(* IEC 61131-3 sources: SRCI_CLIENT_PLC/RobotLibrary/Library/POUs/BasicMove/MC_ReturnToPrimary/Structures, 4 files *)

(* ---- ReturnToPrimaryOutCmd.st ---- *)
{attribute 'pack_mode' := '1'}
// -------------------------------------------------------------------------
//  SRCI Robot Library
// -------------------------------------------------------------------------
//
//  Object:      ReturnToPrimaryOutCmd
//  Author:      Thorsten Brach
//  Date:        2024-06-22
//
//  Description:
//
//
//  Copyright:
//    (C) 2024 Thorsten Brach. All rights reserved
//             Licensed under the MIT License.
//
//  Disclaimer:
//    This project is provided without any guarantee and can be used for
//    private and commercial purposes. Any use is at the user’s
//    own risk and responsibility.
//
// -------------------------------------------------------------------------
TYPE ReturnToPrimaryOutCmd :
STRUCT
  /// Distance-to-go of the current job.
  /// • -1: No valid value because move command is not yet active (valid values are pending) or not supported by RC
  /// • >0: Actual distance between current and target position
  /// •  0: Target position reached
  RemainingDistance  : REAL;
  /// Percentage of already traversed distance of current job.
  /// If not supported : • -1
  Progress           : REAL;
  /// Tool index of target position of ReturnToPrimary
  /// • 0: Flange
  /// • 1..254: Tool frames
  PrimaryPosToolNo   : USINT;
  /// Frame index of target position of ReturnToPrimary
  /// • 0: WCS
  ///• 1..254: User frames
  PrimaryPosFrameNo  : USINT;
END_STRUCT
END_TYPE

(* ---- ReturnToPrimaryParCmd.st ---- *)
{attribute 'pack_mode' := '1'}
// -------------------------------------------------------------------------
//  SRCI Robot Library
// -------------------------------------------------------------------------
//
//  Object:      ReturnToPrimaryParCmd
//  Author:      Thorsten Brach
//  Date:        2024-06-22
//
//  Description:
//
//
//  Copyright:
//    (C) 2024 Thorsten Brach. All rights reserved
//             Licensed under the MIT License.
//
//  Disclaimer:
//    This project is provided without any guarantee and can be used for
//    private and commercial purposes. Any use is at the user’s
//    own risk and responsibility.
//
// -------------------------------------------------------------------------
TYPE ReturnToPrimaryParCmd :
STRUCT
  /// Defines target position when function is executed:
  /// • 0: Interrupt position (default) - Returns to position active,  when interrupt was executed
  /// • 1: End position                 - Returns to target position of interrupted segment
  ReturnMode         : ReturnMode;
  /// TCP velocity in % of nominal velocity
  /// •  <0%: (default) - Use default velocity
  /// •   0%:           - Use internal minimal velocity
  /// • 100%:           - Use maximal reference velocity
  /// See chapter 5.5.7 Robot dynamics
  VelocityRate       : REAL := -1.0; // ST-FIX F41: spec 5.x robot dynamics parameter: '<0 %: use default' (default); the library had 0.0 = internal minimal value (the RC rejects 0 for DecelerationRate/JerkRate)
  /// Acceleration for movement in % of nominal acceleration
  /// •  <0%: (default) - Use default acceleration
  /// •   0%:           - Use internal minimal acceleration
  /// • 100%:           - Use maximal reference acceleration
  /// See chapter 5.5.7 Robot dynamics
  AccelerationRate   : REAL := -1.0; // ST-FIX F41: spec 5.x robot dynamics parameter: '<0 %: use default' (default); the library had 0.0 = internal minimal value (the RC rejects 0 for DecelerationRate/JerkRate)
  /// Deceleration for movement in % of nominal deceleration
  /// •  <0%: (default) - Use default deceleration
  /// •   0%:           - Use internal minimal deceleration
  /// • 100%:           - Use maximal reference deceleration
  /// See chapter 5.5.7 Robot dynamics
  DecelerationRate   : REAL := -1.0; // ST-FIX F41: spec 5.x robot dynamics parameter: '<0 %: use default' (default); the library had 0.0 = internal minimal value (the RC rejects 0 for DecelerationRate/JerkRate)
  /// Jerk of the movement in % of nominal jerk
  /// •  <0%: (default) - Use default jerk
  /// •   0%:           - Use internal minimal jerk
  /// • 100%:           - Use maximal reference jerk
  /// See chapter 5.5.7 Robot dynamics
  JerkRate           : REAL := -1.0; // ST-FIX F41: spec 5.x robot dynamics parameter: '<0 %: use default' (default); the library had 0.0 = internal minimal value (the RC rejects 0 for DecelerationRate/JerkRate)
  /// Index of tool
  /// •      0: Flange (default)
  /// • 1..254: Tool frames
  ToolNo             : USINT;
  /// Index of frame
  /// •      0: WCS (default)
  /// • 1..254: User frames
  FrameNo            : USINT;
  /// Parameter is used if it is greater than 0 (default):
  /// Maximum allowed distance between current position and target position according to ReturnMode.
  /// If calculated distance is beyond specified Limit, RC returns an error
  DistanceLimit      : REAL;
  /// Defines type of command movement. One of the optional modes must be supported
  TrajectoryMode     : TrajectoryMode;
  /// Parameter is used if it is greater than 0 (default)
  /// • Velocity input is ignored
  /// • Parameter defines the time for the movement to reach the target position
  /// Error is sent by the RC if the time cannot be kept
  MoveTime           : TIME;
  /// Set TRUE to deactivate comparison of
  /// • ToolData and FrameData
  /// • ToolNo and PrimaryPosToolNo
  /// • FrameNo and PrimaryPosFrameNo
  AllowDifferences   : BOOL;
END_STRUCT
END_TYPE

(* ---- ReturnToPrimaryRecvData.st ---- *)
{attribute 'pack_mode' := '1'}
// -------------------------------------------------------------------------
//  SRCI Robot Library
// -------------------------------------------------------------------------
//
//  Object:      ReturnToPrimaryRecvData
//  Author:      Thorsten Brach
//  Date:        2024-06-22
//
//  Description:
//
//
//  Copyright:
//    (C) 2024 Thorsten Brach. All rights reserved
//             Licensed under the MIT License.
//
//  Disclaimer:
//    This project is provided without any guarantee and can be used for
//    private and commercial purposes. Any use is at the user’s
//    own risk and responsibility.
//
// -------------------------------------------------------------------------
TYPE ReturnToPrimaryRecvData EXTENDS RspHeader :
STRUCT
  /// Percentage of already traversed distance of current job.
  /// If not supported : • -1
  Progress           : UINT;
  /// Distance-to-go of the current job.
  /// • -1: No valid value because move command is not yet active (valid values are pending) or not supported by RC
  /// • >0: Actual distance between current and target position
  /// •  0: Target position reached
  RemainingDistance  : REAL;
  /// Tool index of target position of ReturnToPrimary
  /// • 0: Flange
  /// • 1..254: Tool frames
  PrimaryPosToolNo   : USINT;
  /// Frame index of target position of ReturnToPrimary
  /// • 0: WCS
  ///• 1..254: User frames
  PrimaryPosFrameNo  : USINT;
END_STRUCT
END_TYPE

(* ---- ReturnToPrimarySendData.st ---- *)
{attribute 'pack_mode' := '1'}
// -------------------------------------------------------------------------
//  SRCI Robot Library
// -------------------------------------------------------------------------
//
//  Object:      ReturnToPrimarySendData
//  Author:      Thorsten Brach
//  Date:        2024-06-22
//
//  Description:
//
//
//  Copyright:
//    (C) 2024 Thorsten Brach. All rights reserved
//             Licensed under the MIT License.
//
//  Disclaimer:
//    This project is provided without any guarantee and can be used for
//    private and commercial purposes. Any use is at the user’s
//    own risk and responsibility.
//
// -------------------------------------------------------------------------
TYPE ReturnToPrimarySendData EXTENDS CmdHeader:
STRUCT
  /// TCP velocity in % of nominal velocity
  /// •  <0%: (default) - Use default velocity
  /// •   0%:           - Use internal minimal velocity
  /// • 100%:           - Use maximal reference velocity
  /// See chapter 5.5.7 Robot dynamics
  VelocityRate       : UINT;
  /// Acceleration for movement in % of nominal acceleration
  /// •  <0%: (default) - Use default acceleration
  /// •   0%:           - Use internal minimal acceleration
  /// • 100%:           - Use maximal reference acceleration
  /// See chapter 5.5.7 Robot dynamics
  AccelerationRate   : UINT;
  /// Deceleration for movement in % of nominal deceleration
  /// •  <0%: (default) - Use default deceleration
  /// •   0%:           - Use internal minimal deceleration
  /// • 100%:           - Use maximal reference deceleration
  /// See chapter 5.5.7 Robot dynamics
  DecelerationRate   : UINT;
  /// Jerk of the movement in % of nominal jerk
  /// •  <0%: (default) - Use default jerk
  /// •   0%:           - Use internal minimal jerk
  /// • 100%:           - Use maximal reference jerk
  /// See chapter 5.5.7 Robot dynamics
  JerkRate           : UINT;
  /// Parameter is used if it is greater than 0 (default):
  /// Maximum allowed distance between current position and target position according to ReturnMode.
  /// If calculated distance is beyond specified Limit, RC returns an error
  DistanceLimit      : REAL;
  /// Index of tool
  /// •      0: Flange (default)
  /// • 1..254: Tool frames
  ToolNo             : USINT;
  /// Index of frame
  /// •      0: WCS (default)
  /// • 1..254: User frames
  FrameNo            : USINT;
  /// Parameter is used if it is greater than 0 (default)
  /// • Velocity input is ignored
  /// • Parameter defines the time for the movement to reach the target position
  /// Error is sent by the RC if the time cannot be kept
  MoveTime           : UINT;
  /// Defines target position when function is executed:
  /// • 0: Interrupt position (default) - Returns to position active,  when interrupt was executed
  /// • 1: End position                 - Returns to target position of interrupted segment
  ReturnMode         : BOOL;
  /// Defines type of command movement. One of the optional modes must be supported
  TrajectoryMode     : BOOL;
  ///
  Enable : BOOL;
  ///
  AllowDifferences : BOOL;

END_STRUCT
END_TYPE
